FUNCTION FC 1 : VOID
BEGIN
NETWORK
      BE 1
END_FUNCTION
